// TIA Portal V20 export
TYPE "DataRange"
   STRUCT
      inRange : Array[0..2000] of Byte;
   END_STRUCT;
END_TYPE
